// TIA Portal V20 export
// export: Created 2026-10-19T18:44:24.3603179Z, ExportSetting WithDefaults, DisplayName Totally Integrated Automation Portal, DisplayVersion V20 Update 6, DisplayName TIA Portal Openness, DisplayVersion V20 Update 6, DisplayName TIA Portal Version Control Interface, DisplayVersion V20 Update 6, DisplayName SINAMICS Startdrive Advanced, DisplayVersion V20 SP1, DisplayName SINAMICS Startdrive G130, G150, S120, S150, SINAMICS MV, G220, S200, S210, DisplayVersion V20 SP1, DisplayName SINAMICS Startdrive G110M, G120, G120C, G120D, G120P, G115D, DisplayVersion V20 SP1, DisplayName STEP 7 Professional, DisplayVersion V20 Update 6, DisplayName STEP 7 Safety, DisplayVersion V20 Update 2, DisplayName WinCC Basic/Comfort/Advanced, DisplayVersion V20 Update 6, DisplayName WinCC Unified, DisplayVersion V20 Update 6
DATA_BLOCK "LCom_Comm_Shuttle_FB_DB_10"   // DB359
AUTHOR : APC_ERLF
FAMILY : LCom
VERSION : 2.1
// stored: AutoNumber true, DBAccessibleFromOPCUA true, InstanceOfName LCom_Communication_FB, InstanceOfType FB
"LCom_Communication_FB"
   // VAR_INPUT
   //    enable : Bool;
   //    send : Bool;
   //    sendDataLength : UDInt;
   //    readDataLength : UDInt;
   //    configuration : "LCom_typeConfig";
   // END_VAR
   // VAR_OUTPUT
   //    connected : Bool;
   //    sending : Bool;
   //    dataReceived : Bool;
   //    receivedDataLength : UDInt;
   //    busy : Bool;
   //    error : Bool;
   //    status : Word;
   // END_VAR
   // VAR_IN_OUT
   //    sendBuffer : Variant;
   //    receiveBuffer : Variant;
   //    diagnostics : "LCom_typeDiagnostics";
   // END_VAR
   // VAR
   //    statConnectAttempts : SInt;
   //    statActualLocalLComVersion : USInt;
   //    statRuntimeTask : LReal;
   //    statCopyNBytes : UDInt;
   //    statMaxActPacketLength : UDInt;
   //    statState : Struct
   //       connection : USInt;
   //       cfgSender : USInt;
   //       comSender : USInt;
   //       comReceiver : USInt;
   //       sender : USInt;
   //       receiver : USInt;
   //    END_STRUCT;
   //    statReceive : Struct
   //       tempTelegram : Struct
   //          LComVersion : USInt;
   //          index : USInt;
   //          telegramType : USInt;
   //          data : Array[0..23] of Byte;
   //       END_STRUCT;
   //       configTelegramV1 : Struct
   //          LComVersion : USInt;
   //          telegramType : USInt;
   //          comMode : USInt;
   //          slidingWindow : USInt;
   //          cycleTime : UInt;
   //          ackTimeOut : UInt;
   //          lifeSignCycle : UInt;
   //          status : USInt;
   //          sendModeSyncTime : USInt;
   //          maxSendDataLength : UInt;
   //          maxReceiveDataLength : UInt;
   //       END_STRUCT;
   //       configTelegramV2 : Struct
   //          LComVersion : USInt;
   //          telegramType : USInt;
   //          status : USInt;
   //          sendModeSyncTime : USInt;
   //          lifeSignCycle : Time;
   //          cycleTime : Time;
   //          ackTimeOut : Time;
   //          maxSendDataLength : UDInt;
   //          maxReceiveDataLength : UDInt;
   //       END_STRUCT;
   //       dataTelegram : Struct
   //          LComVersion : USInt;
   //          telegramType : USInt;
   //          messageCounter : USInt;
   //          ackMessageCounter : USInt;
   //          messageOffset : UDInt;
   //          ackMessageOffset : UDInt;
   //          actPackageLength : UDInt;
   //          totalMessageLength : UDInt;
   //       END_STRUCT;
   //       userData : Struct
   //          totalLength : UDInt;
   //          offset : UDInt;
   //       END_STRUCT;
   //       trcvFct : Struct
   //          data : Array[0..4095] of Byte;
   //          dataOffset : UDInt;
   //          dataLength : UDInt;
   //          dataLengthRest : UDInt;
   //          dataReceived : Bool;
   //       END_STRUCT;
   //       numberOfLComHeader : USInt;
   //    END_STRUCT;
   //    statSend : Struct
   //       configTelegramV1 : Struct
   //          LComVersion : USInt;
   //          comMode : USInt;
   //          slidingWindow : USInt;
   //          cycleTime : UInt;
   //          ackTimeOut : UInt;
   //          lifeSignCycle : UInt;
   //          status : USInt;
   //          sendModeSyncTime : USInt;
   //          maxSendDataLength : UInt;
   //          maxReceiveDataLength : UInt;
   //       END_STRUCT;
   //       configTelegramV2 : Struct
   //          LComVersion : USInt;
   //          status : USInt;
   //          sendModeSyncTime : USInt;
   //          lifeSignCycle : Time;
   //          cycleTime : Time;
   //          ackTimeOut : Time;
   //          maxSendDataLength : UDInt;
   //          maxReceiveDataLength : UDInt;
   //       END_STRUCT;
   //       dataTelegram : Struct
   //          LComVersion : USInt;
   //          telegramType : USInt;
   //          messageCounter : USInt;
   //          ackMessageCounter : USInt;
   //          messageOffset : UDInt;
   //          ackMessageOffset : UDInt;
   //          actPackageLength : UDInt;
   //          totalMessageLength : UDInt;
   //       END_STRUCT;
   //       userData : Struct
   //          totalLength : UDInt;
   //          offset : UDInt;
   //          sendCycleViolation : Bool;
   //       END_STRUCT;
   //       tsendFct : Struct
   //          dataLengthRest : UInt;
   //          data : Array[0..4095] of Byte;
   //          dataOffset : UInt;
   //          status : Word;
   //          enable : Bool;
   //       END_STRUCT;
   //       expectedAck : Struct
   //          package1 : Struct
   //             offset : UDInt;
   //          END_STRUCT;
   //       END_STRUCT;
   //       numberOfLComPackage : USInt;
   //    END_STRUCT;
   //    statIterator : Int;
   //    statOldEnable : Bool;
   //    statOldSend : Bool;
   //    statRisingEdgeSend : Bool;
   //    statFallingEdgeEnable : Bool;
   //    statRet : Int;
   //    statCompare : Struct
   //       sender : Struct
   //          cycleTime : Time;
   //          ackTimeOut : Time;
   //       END_STRUCT;
   //    END_STRUCT;
   //    statTconPar { S7_SetPoint := 'True'} : TCON_IP_v4;
   //    statTconParQdn { S7_SetPoint := 'True'} : TCON_QDN;
   //    instTCON { S7_SetPoint := 'True'} : TCON;
   //    instTDISCON { S7_SetPoint := 'True'} : TDISCON;
   //    instTRCV { S7_SetPoint := 'True'} : TRCV;
   //    instTSEND { S7_SetPoint := 'True'} : TSEND;
   //    instLocalLifeSignCycleTimer { S7_SetPoint := 'True'} : TON_TIME;
   //    instPartnerLifeSignCycleTimer { S7_SetPoint := 'True'} : TON_TIME;
   //    instLocalCycleTimeTimer { S7_SetPoint := 'True'} : TON_TIME;
   //    instReceiveMsgCycle { S7_SetPoint := 'True'} : TON_TIME;
   //    instExpectedAckPackage1 { S7_SetPoint := 'True'} : TON_TIME;
   //    instMsgSendingTimer { S7_SetPoint := 'True'} : TON_TIME;
   //    instMsgReceivingTimer { S7_SetPoint := 'True'} : TON_TIME;
   //    instSyncTimer { S7_SetPoint := 'True'} : TON_TIME;
   //    instSendErrorTimer { S7_SetPoint := 'True'} : TON_TIME;
   //    instRcvErrorTimer { S7_SetPoint := 'True'} : TON_TIME;
   //    instRDREC { S7_SetPoint := 'True'} : RDREC;
   //    statDiag : Struct
   //       buffer : Array[0..9] of Struct
   //          status : Word;
   //          isActive : Bool;
   //          subFunctionErrorID : Word;
   //          additionalValue1 : Real;
   //          additionalValue2 : Real;
   //          additionalValue3 : Real;
   //          additionalValue4 : Time;
   //       END_STRUCT;
   //       bufferIndex : Int;
   //       actualIndex : USInt;
   //    END_STRUCT;
   //    statDataReceived : Bool;
   //    statConnected : Bool;
   //    statStatus : Word;
   //    statSending : Bool;
   // END_VAR
BEGIN
END_DATA_BLOCK
